(* PLC project Vn_sub, Beckhoff Automation GmbH TwinCAT PLC Control 3.5.13.21 *)
(* stored: creationDateTime 1970-01-01T00:00:00 *)

PROGRAM Vn_sub

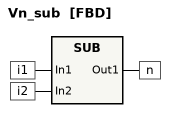
(* FBD diagram, written out as Structured Text *)
n := i1 - i2;
END_PROGRAM
